FUNCTION_BLOCK TestingStation (* Composite Function Block Type *)
  (* Standard: 61499-2 *)
  (* Version 0.0, 7/2/2026, template *)
  PACKAGE Main;
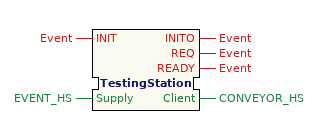
  EVENT_INPUT
    INIT; (* Initialization Request *)
  END_EVENT
  EVENT_OUTPUT
    INITO; (* Initialization Confirm *)
    REQ; (* Execution Confirmation *)
    READY;
  END_EVENT
  SOCKETS
    Supply : EVENT_HS;
  END_SOCKETS
  PLUGS
    Client : CONVEYOR_HS;
  END_PLUGS
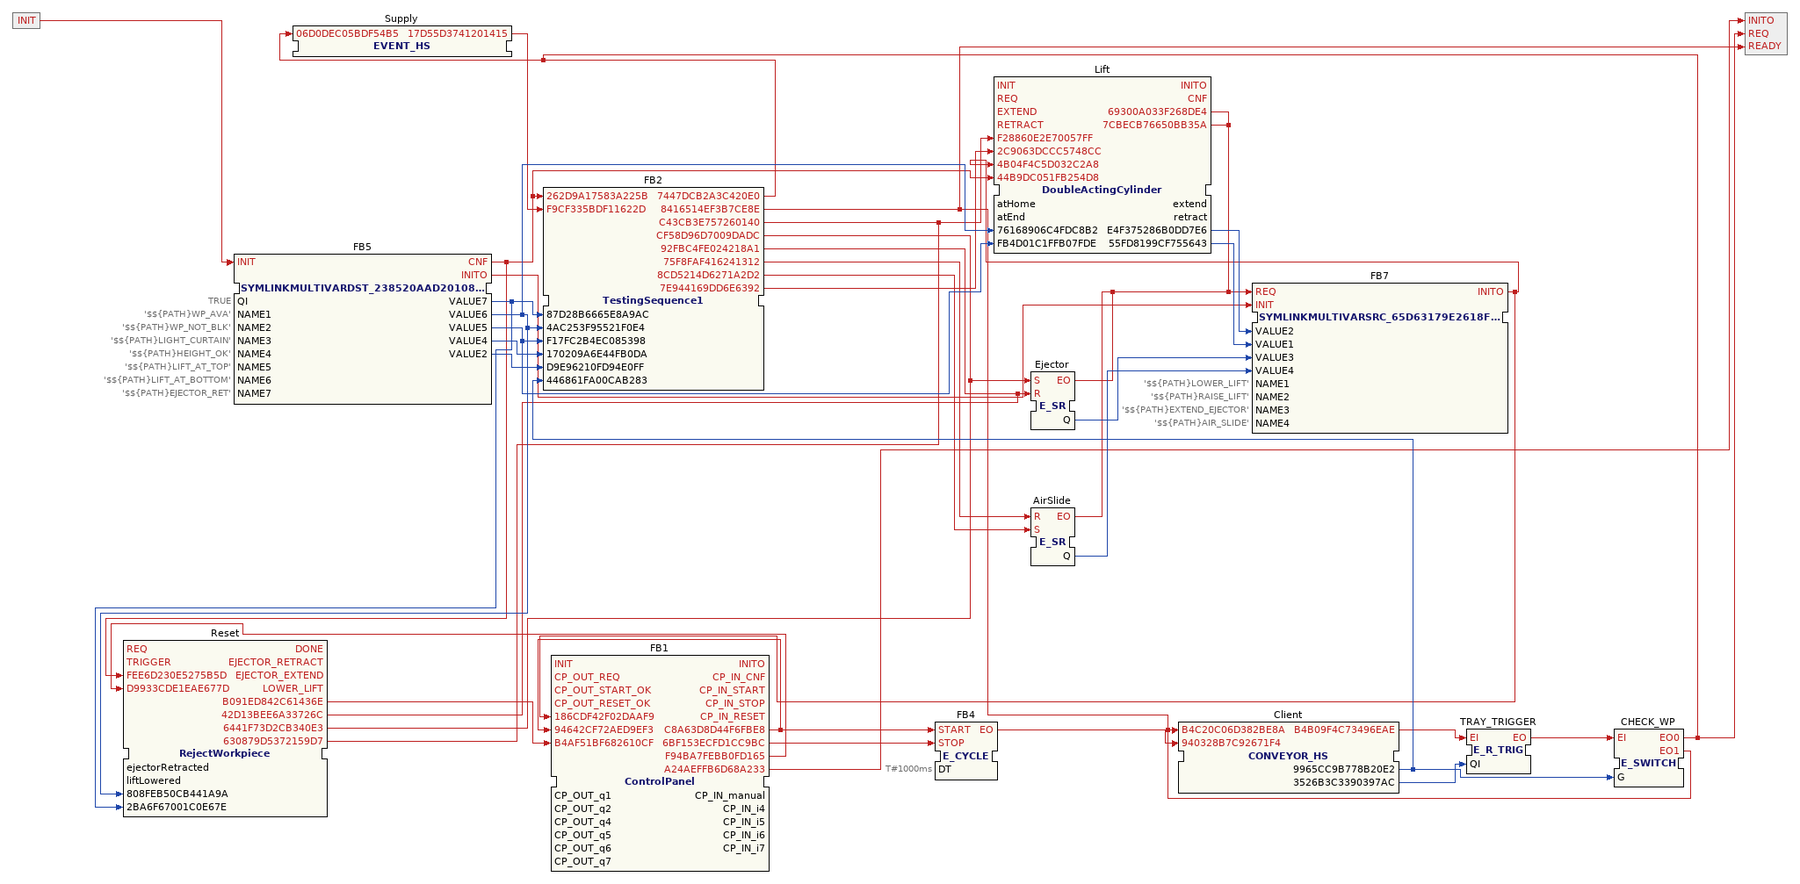
  FBS
    FB2 : TestingSequence1;
    FB5 : SYMLINKMULTIVARDST_238520AAD20108C65(QI := TRUE, NAME1 := '$${PATH}WP_AVA', NAME2 := '$${PATH}WP_NOT_BLK', NAME3 := '$${PATH}LIGHT_CURTAIN', NAME4 := '$${PATH}HEIGHT_OK', NAME5 := '$${PATH}LIFT_AT_TOP', NAME6 := '$${PATH}LIFT_AT_BOTTOM', NAME7 := '$${PATH}EJECTOR_RET'); {SET_ATTRIBUTE(Configuration.GenericFBType.InterfaceParams, Runtime.System#I:=7;VALUE${I$}:BOOL,BOOL,BOOL,BOOL,BOOL,BOOL,BOOL)}
    FB7 : SYMLINKMULTIVARSRC_65D63179E2618F5E(NAME1 := '$${PATH}LOWER_LIFT', NAME2 := '$${PATH}RAISE_LIFT', NAME3 := '$${PATH}EXTEND_EJECTOR', NAME4 := '$${PATH}AIR_SLIDE'); {SET_ATTRIBUTE(Configuration.GenericFBType.InterfaceParams, Runtime.System#I:=5;VALUE${I$}:BOOL,BOOL,BOOL,BOOL,BOOL)}
    Lift : DoubleActingCylinder;
    Ejector : E_SR;
    AirSlide : E_SR;
    FB4 : E_CYCLE(DT := T#1000ms);
    TRAY_TRIGGER : E_R_TRIG;
    CHECK_WP : E_SWITCH;
    FB1 : ControlPanel;
    Reset : RejectWorkpiece;
  END_FBS
  EVENT_CONNECTIONS
    INIT TO FB5.INIT;
    FB5.CNF TO FB2.262D9A17583A225B;
    Supply.17D55D3741201415 TO FB2.F9CF335BDF11622D;
    FB2.7447DCB2A3C420E0 TO Supply.06D0DEC05BDF54B5;
    CHECK_WP.EO0 TO Supply.06D0DEC05BDF54B5;
    FB2.8416514EF3B7CE8E TO READY;
    FB2.8416514EF3B7CE8E TO Client.B4C20C06D382BE8A;
    FB2.C43CB3E757260140 TO Lift.F28860E2E70057FF;
    FB2.CF58D96D7009DADC TO Ejector.S;
    FB2.92FBC4FE024218A1 TO Ejector.R;
    FB2.75F8FAF416241312 TO AirSlide.R;
    FB2.8CD5214D6271A2D2 TO AirSlide.S;
    FB2.7E944169DD6E6392 TO Lift.2C9063DCCC5748CC;
    Lift.69300A033F268DE4 TO FB7.REQ;
    Lift.7CBECB76650BB35A TO FB7.REQ;
    Ejector.EO TO FB7.REQ;
    AirSlide.EO TO FB7.REQ;
    FB7.INITO TO Lift.4B04F4C5D032C2A8;
    FB7.INITO TO FB1.186CDF42F02DAAF9;
    FB5.CNF TO Lift.44B9DC051FB254D8;
    FB5.CNF TO Reset.FEE6D230E5275B5D;
    FB5.INITO TO FB7.INIT;
    CHECK_WP.EO0 TO REQ;
    CHECK_WP.EO1 TO Client.B4C20C06D382BE8A;
    TRAY_TRIGGER.EO TO CHECK_WP.EI;
    Client.B4B09F4C73496EAE TO TRAY_TRIGGER.EI;
    FB4.EO TO Client.940328B7C92671F4;
    FB1.C8A63D8D44F6FBE8 TO FB4.START;
    FB1.6BF153ECFD1CC9BC TO FB4.STOP;
    FB1.C8A63D8D44F6FBE8 TO FB1.94642CF72AED9EF3;
    Reset.B091ED842C61436E TO FB1.B4AF51BF682610CF;
    FB1.F94BA7FEBB0FD165 TO Reset.D9933CDE1EAE677D;
    FB1.A24AEFFB6D68A233 TO INITO;
    Reset.42D13BEE6A33726C TO Ejector.R;
    Reset.6441F73D2CB340E3 TO Ejector.S;
    Reset.630879D5372159D7 TO Lift.F28860E2E70057FF;
  END_CONNECTIONS
  DATA_CONNECTIONS
    FB5.VALUE7 TO FB2.87D28B6665E8A9AC;
    FB5.VALUE6 TO FB2.4AC253F95521F0E4;
    FB5.VALUE5 TO FB2.F17FC2B4EC085398;
    FB5.VALUE4 TO FB2.170209A6E44FB0DA;
    FB5.VALUE2 TO FB2.D9E96210FD94E0FF;
    Client.9965CC9B778B20E2 TO FB2.446861FA00CAB283;
    FB5.VALUE6 TO Lift.76168906C4FDC8B2;
    FB5.VALUE5 TO Lift.FB4D01C1FFB07FDE;
    Lift.E4F375286B0DD7E6 TO FB7.VALUE2;
    Lift.55FD8199CF755643 TO FB7.VALUE1;
    Ejector.Q TO FB7.VALUE3;
    AirSlide.Q TO FB7.VALUE4;
    Client.9965CC9B778B20E2 TO CHECK_WP.G;
    Client.3526B3C3390397AC TO TRAY_TRIGGER.QI;
    FB5.VALUE6 TO Reset.808FEB50CB441A9A;
    FB5.VALUE7 TO Reset.2BA6F67001C0E67E;
  END_CONNECTIONS
END_FUNCTION_BLOCK
